Fanuc KAREL source: KB00137.KL

PROGRAM KB00137
%NOLOCKGROUP
%ENVIRONMENT CORE
VAR
  P1: STRING[80]
  P2: INTEGER
  P3: INTEGER
  P4: BOOLEAN
  P5: INTEGER
BEGIN
  P1 = 'A'
  P2 = 1
  P3 = 1
  P4 = TRUE
  P5 = 1
  PROG_BACKUP(P1, P2, P3, P4, P5)
END KB00137
